Staubli VAL3: kill.pgx

public program kill()
begin
  //Kill Task
  taskKill("actCtrl")
  wait(taskStatus("actCtrl")==-1)
  call clearActStack()
end
